// TIA Portal V21 export
FUNCTION "FC_FbdLogic" : Void   // FC8, FBD
TITLE = FUP-Logik / FBD logic
{ S7_Optimized_Access := 'TRUE' }
// UND, ODER, XOR, Negation, Zuweisung, SR, RS und Flankenerkennung in FUP / AND, OR, XOR, negation, assignment, SR, RS and edge detection in FBD
// stored: SetENOAutomatically false
   VAR_INPUT
      InA : Bool;
      InB : Bool;
   END_VAR
   VAR_OUTPUT
      AndOut : Bool;
      OrOut : Bool;
      XorOut : Bool;
      NotOut : Bool;
      SrOut : Bool;
      RsOut : Bool;
      EdgeOut : Bool;
   END_VAR
   VAR_IN_OUT
      SrBit : Bool;
      RsBit : Bool;
      EdgeBit : Bool;
   END_VAR
   VAR_TEMP   // added for the SCL form of the ladder/FBD networks
      _w1 : Bool;
   END_VAR
BEGIN

REGION Network 1: UND / AND
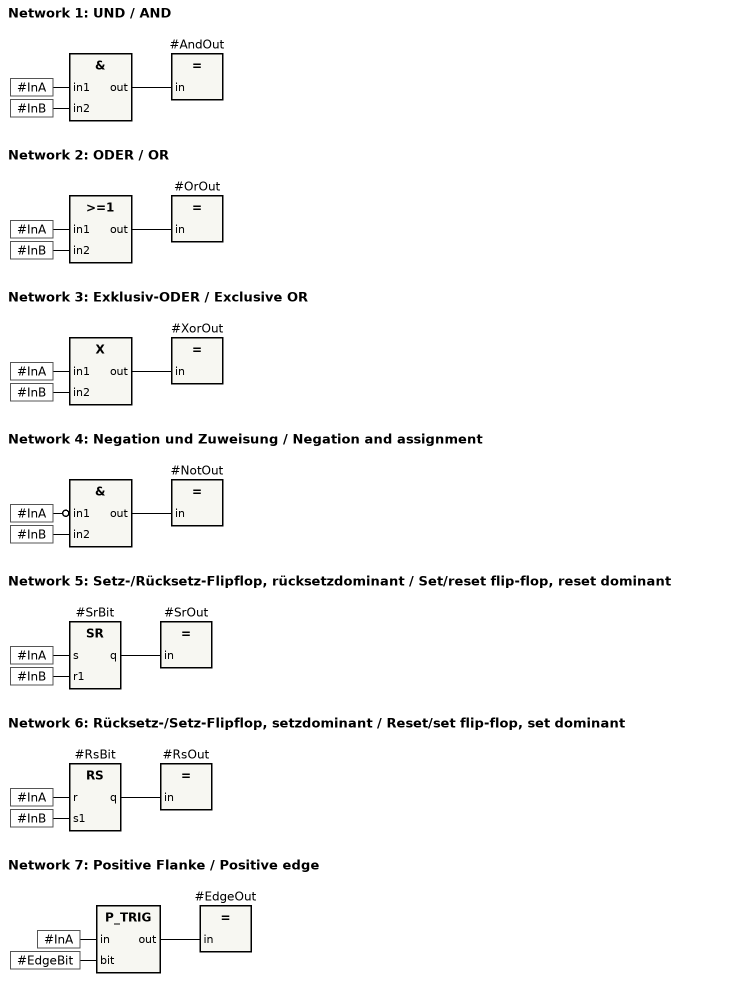
   #AndOut := #InA AND #InB;
END_REGION

REGION Network 2: ODER / OR
   #OrOut := #InA OR #InB;
END_REGION

REGION Network 3: Exklusiv-ODER / Exclusive OR
   #XorOut := #InA XOR #InB;
END_REGION

REGION Network 4: Negation und Zuweisung / Negation and assignment
   #NotOut := NOT #InA AND #InB;
END_REGION

REGION Network 5: Setz-/Rücksetz-Flipflop, rücksetzdominant / Set/reset flip-flop, reset dominant
   IF #InA THEN
       #SrBit := TRUE;   // SR flip-flop
   END_IF;
   IF #InB THEN #SrBit := FALSE; END_IF;
   #SrOut := #SrBit;
END_REGION

REGION Network 6: Rücksetz-/Setz-Flipflop, setzdominant / Reset/set flip-flop, set dominant
   IF #InA THEN
       #RsBit := FALSE;   // RS flip-flop
   END_IF;
   IF #InB THEN #RsBit := TRUE; END_IF;
   #RsOut := #RsBit;
END_REGION

REGION Network 7: Positive Flanke / Positive edge
   #_w1 := #InA AND NOT #EdgeBit;   // rising edge
   #EdgeBit := #InA;
   #EdgeOut := #_w1;
END_REGION
END_FUNCTION
